Fanuc KAREL source: KA00015.KL

PROGRAM KA00015
%NOLOCKGROUP
VAR
  SRC: REAL
  DST: BOOLEAN
BEGIN
  SRC = 2.0
  DST = SRC
END KA00015
